// TIA Portal V20 export
FUNCTION "Real Laden" : Void   // FC131, STL
TITLE = Real Laden für Graph
{ S7_Optimized_Access := 'FALSE' }
// stored: AutoNumber false
   VAR_INPUT
      Eingabewert : Real;
   END_VAR
   VAR_OUTPUT
      Ausgabewert : Real;
   END_VAR
BEGIN

NETWORK
TITLE = 
      L     #Eingabewert;
      T     #Ausgabewert;
END_FUNCTION
